// TIA Portal V21 export
TextList "TL_Alarm"  ListRange=Decimal
  TextListEntry   From=-1, To=-1, Text="-"
  TextListEntry   Text="0 Neuravnoteženost broda |L-R| > 5"
  TextListEntry   From=1, To=1, Text="1 Lokacija podizanja prazna"
  TextListEntry   From=2, To=2, Text="2 Lokacija spuštanja zauzeta"
  TextListEntry   From=3, To=3, Text="3 ID kontejnera postoji u listi za istovar, ali ne postoji u polju Bay 0"
  TextListEntry   From=4, To=4, Text="4 ID kontejnera postoji u listi za ukrcaj, ali ne postoji u polju Bay 1"
  TextListEntry   From=5, To=5, Text="5 Neispravan ID (100-999)"
  TextListEntry   From=6, To=6, Text="6 Dvostruki ID"
  TextListEntry   From=7, To=7, Text="7 Nema slobodnog mjesta"
  TextListEntry   From=8, To=8, Text="8 Plan nije izvediv"
  TextListEntry   From=9, To=9, Text="9 Neispravna ručna naredba"
  TextListEntry   From=10, To=10, Text="10 Dizalica: timeout naredbe"
  TextListEntry   From=11, To=11, Text="11 Dizalica već nosi kontejner"
  TextListEntry   From=12, To=12, Text="12 Dizalica ne nosi kontejner"
  TextListEntry   From=13, To=13, Text="13 Nije inicijalizirano"
  TextListEntry   From=14, To=14, Text="14 Položaj dizalice ne odgovara"
  TextListEntry   From=15, To=15, Text="15 Istovar i ukrcaj završeni"
